FUNCTION_BLOCK MOD_OwnerLatch (* Keeps the last owner heard on the owner channel. Technical: Local channel IDs of the occupation owner and its refresh query; types and forwards the received occupation owner *)
  (* Standard: 61499-2 *)
  (* Version 0.1, 2026-09-28, Project contributors, AAU Smart Production Lab *)
  PACKAGE modlib;
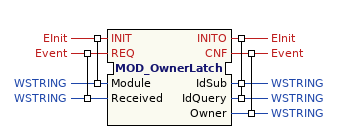
  EVENT_INPUT
    INIT : EInit WITH Module; (* Initialise, once at start-up (the INIT chain); takes the values given with it *)
    REQ WITH Received; (* The value arrived on the local channel *)
  END_EVENT
  EVENT_OUTPUT
    INITO : EInit WITH IdSub, IdQuery; (* Initialised: the next block of the INIT chain goes on *)
    CNF WITH Owner; (* Confirmation of REQ *)
  END_EVENT
  VAR_INPUT
    Module : WSTRING; (* The module's name; its local channels are named after it (loc[<Module>/...]) *)
    Received : WSTRING; (* The value as it arrived *)
  END_VAR
  VAR_OUTPUT
    IdSub : WSTRING; (* Local channel the value arrives on *)
    IdQuery : WSTRING; (* Local channel that asks for the current value (a block that starts later) *)
    Owner : WSTRING; (* Session ID of the module's owner (empty: free) *)
  END_VAR
  EC_STATES
    INIT : INIT -> INITO;
    REQ : REQ -> CNF;
  END_STATES
  ALGORITHM INIT IN ST:
IdSub := CONCAT(CONCAT("loc[", Module), "/owner]");
IdQuery := CONCAT(CONCAT("loc[", Module), "/owner/query]");
  END_ALGORITHM
  ALGORITHM REQ IN ST:
Owner := Received;
  END_ALGORITHM
END_FUNCTION_BLOCK
